Fanuc KAREL source: kb00037.KL

-- PROVISIONAL review KL for V770-1; original PC SHA256 16a2ec077f4bb63c4873c2babaf23b4aaaaf3afe436376e43117809d2df40293
-- Incomplete behavior may be omitted. Consult companion uncertainty JSON. Do not deploy.
PROGRAM KB00037
%NOLOCKGROUP
BEGIN
  -- UNRESOLVED_PC offsets 5-16; opcodes 2E,23
  -- UNRESOLVED_PC offsets 21-28; opcodes 9D,23
  -- UNRESOLVED_PC offsets 33-40; opcodes 9D,23
  -- UNRESOLVED_PC offsets 45-54; opcodes 3F,75
  -- UNRESOLVED_PC offsets 59-89; opcodes 27,22,22,22,22,2A,31
  -- UNRESOLVED_PC offsets 94-98; opcodes 7F
END KB00037
